Universal Robots PolyScope program: PgProg.urp

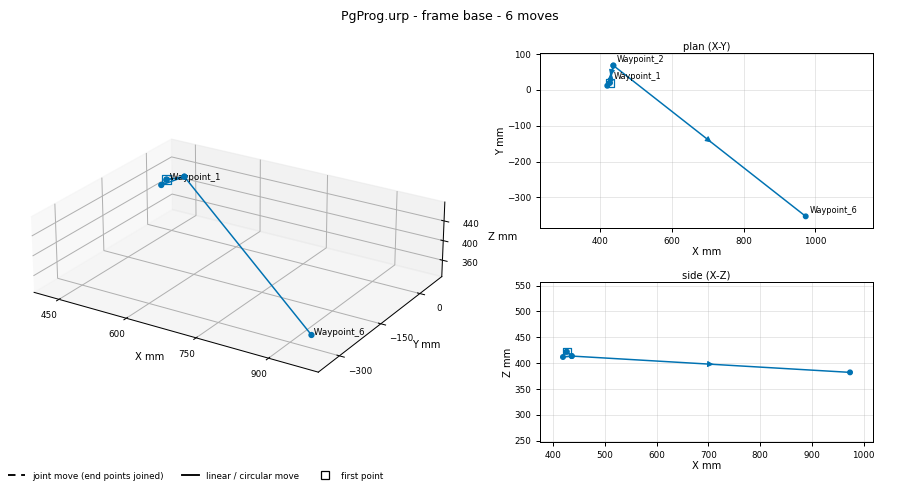
[picture p0: tool path of PgProg.urp in frame base, 6 of 6 moves have a stored position in this frame; points joined in program order, loops and branches not executed]
Program PgProg (createdIn=3.0.0 lastSavedIn=3.0.0 directory=/programs installation=default)
Robot Program (runOnlyOnce=true motionType=MoveJ speed=1.047198 acceleration=1.396263 useActiveTCP=false)
  'Program generated by RoboDK v6.0.7 for ABB IRB 120-3/0.6 on XX/XX/XXXX 18:00:00'
  'Using nominal kinematics.'
  'Using Ref. Frame Pg: p[1.234570, -0.098765, 0.050500, 0.000000, 0.000000, 0.523599]'
  'Using TCP Tool Pg: p[0.010000, 0.020000, 0.150000, 0.261799, 0.000000, 0.000000]'
  Script: set_tcp(p[0.010000, 0.020000, 0.150000, 0.261799, 0.000000, 0.000000])
  Script: movej([0.000000, -0.174533, 0.349066, 0.000000, 0.523599, 0.000000],1.20000,0.75000,0,0.0000)
  MoveJ speed 42.97 deg/s, acceleration 68.75 deg/s^2 (useActiveTCP=true)
    Waypoint Waypoint_1: TCP in base x=426.318 y=20 z=422.034 mm, rx=0.1383 ry=2.2532 rz=-0.2966 rad; joints [0, -10, 20, 0, 30, 0] deg; flange x=317.839 y=0 z=526.113 mm, rx=0 ry=2.2689 rz=0 rad
  MoveL speed 250 mm/s, acceleration 1200 mm/s^2 (useActiveTCP=true)
    Waypoint Waypoint_2: motionParameters(blendRadius=0.005); TCP in base x=436.232 y=68.297 z=413.715 mm, rx=0.1383 ry=2.2532 rz=-0.2966 rad; joints [0, -10, 20, 0, 30, 0] deg; flange x=327.753 y=48.297 z=517.794 mm, rx=0 ry=2.2689 rz=0 rad
  'Circular move (R50.0 mm)'
  Script: movec(p[0.414005, 0.116593, 0.367095, 0.138328, 2.253250, -0.296646],p[0.371953, 0.068296, 0.337111, 0.138328, 2.253250, -0.296646],1.20000,0.25000,0.0050)
  Script: movej([0.349066, -0.174533, 0.349066, 0.000000, 0.523599, 0.000000],1.20000,0.75000,0,0.0000)
  MoveL speed 100 mm/s, acceleration 800 mm/s^2 (useActiveTCP=true)
    Waypoint Waypoint_3: motionParameters(blendRadius=0.005); TCP in base x=419.189 y=11.793 z=411.899 mm, rx=0.1383 ry=2.2532 rz=-0.2966 rad; joints [0, -10, 20, 0, 30, 0] deg; flange x=310.711 y=-8.207 z=515.978 mm, rx=0 ry=2.2689 rz=0 rad
    Waypoint Waypoint_4: TCP in base x=426.318 y=20 z=422.034 mm, rx=0.1383 ry=2.2532 rz=-0.2966 rad; joints [0, -10, 20, 0, 30, 0] deg; flange x=317.839 y=0 z=526.113 mm, rx=0 ry=2.2689 rz=0 rad
  Wait Sleep waitTime=0.5
  Halt
  Popup Message (haltProgram=false message=Hello from postgen)
  'a comment'
  Call SubProgram
  Script: CustomCode(42)
  Script: ThreadProg
  Set DigitalOutput pin=digital_out[1]; digitalValue=1
  Set DigitalOutput pin=Valve; digitalValue=0
  Set DigitalOutput pin=digital_out[3]; digitalValue=2.5
  Wait DigitalInput pin=digital_in[get_standard_digital_in(2)]; digitalValue=1
  Wait DigitalInput pin=digital_in[get_standard_digital_in(4)]; digitalValue=0
  'Using TCP Tool2: p[0.000000, 0.000000, 0.200000, 0.000000, 0.000000, 0.000000]'
  Script: set_tcp(p[0.000000, 0.000000, 0.200000, 0.000000, 0.000000, 0.000000])
  Script: movej([0.000000, -0.174533, 0.349066, 0.000000, 0.523599, 0.000000],2.09440,1.04720,0,0.0000)
  MoveJ speed 59.99 deg/s, acceleration 119.98 deg/s^2 (useActiveTCP=true)
    Waypoint Waypoint_5: TCP in base x=436.232 y=68.297 z=413.715 mm, rx=0.1383 ry=2.2532 rz=-0.2966 rad; joints [0, -10, 20, 0, 30, 0] deg; flange x=288.244 y=120.06 z=537.892 mm, rx=0.1383 ry=2.2532 rz=-0.2966 rad
  Script: movej([0.174533, -0.087266, 0.436332, 0.087266, 0.610865, 0.087266],2.09440,1.04720,0,0.0000)
  MoveL speed 100 mm/s, acceleration 800 mm/s^2 (useActiveTCP=true)
    Waypoint Waypoint_6: TCP in base x=973.908 y=-353.337 z=382.202 mm, rx=-0.5037 ry=2.3595 rz=0.0001 rad; joints [-5, -5, 15, 10, 40, -10] deg; flange x=843.629 y=-381.169 z=531.376 mm, rx=-0.5037 ry=2.3595 rz=0.0001 rad
SubProgram  [hidden by the author, left out]
SubProgram SubProgram [hidden by the author, left out]
